Fanuc KAREL source: ko00096.KL

-- PROVISIONAL review KL for V770-1; original PC SHA256 12eebaea0c5418f4bc5985bd2d6ddcee6c8aba9aec44a7e6fc8fe47d6110594f
-- Incomplete behavior may be omitted. Consult companion uncertainty JSON. Do not deploy.
PROGRAM KO00096
%NOLOCKGROUP
BEGIN
  -- UNRESOLVED_PC offsets 5-12; opcodes 9D,23
  -- UNRESOLVED_PC offsets 17-69; opcodes 27,27,49,7E,AD,27,49,7E,AD,22,31,7E,4A
  -- UNRESOLVED_PC offsets 74-78; opcodes 7F
END KO00096
